{region 'Documentation'}
(*!
<summary>Check that IN is inside the inclusive StartTime..EndTime interval.</summary>
<description>

StartTime &gt; EndTime reports Error during active evaluation; equal bounds are
valid.

A value at or beyond 24 hours reports Error before comparison or baseline capture.

</description>
*)
{endregion}
FUNCTION_BLOCK AssertInTimespan_TOD EXTENDS AssertionBase
VAR_INPUT
    IN : TOD; //! Actual value checked or observed by this Assertion.
    StartTime : TOD; //! Inclusive start of the time span; must not exceed EndTime.
    EndTime : TOD; //! Inclusive end of the time span; must not precede StartTime.
END_VAR

SUPER^();

{region 'Documentation'}
(*!
<summary>Evaluate the typed temporal relation and report higher-priority errors first.</summary>
*)
{endregion}
METHOD PROTECTED Assert
VAR
    Message : STRING(GVL_Constants.MessageLength);
    StartTimeText : STRING(GVL_Constants.AssertionValueLength);
    EndTimeText : STRING(GVL_Constants.AssertionValueLength);
    ActualText : STRING(GVL_Constants.AssertionValueLength);
END_VAR
IF NOT EvaluationActive THEN
    RETURN;
END_IF;

IF Result = E_Result.Error THEN
    RETURN;
END_IF;

IF NOT IsTimeOfDayValid_TOD(Value := IN) THEN
    Error(Message := 'Assertion error: IN is outside the valid TOD range (less than 24 hours).');
    RETURN;
END_IF;

IF NOT IsTimeOfDayValid_TOD(Value := StartTime) THEN
    Error(Message := 'Assertion error: StartTime is outside the valid TOD range (less than 24 hours).');
    RETURN;
END_IF;

IF NOT IsTimeOfDayValid_TOD(Value := EndTime) THEN
    Error(Message := 'Assertion error: EndTime is outside the valid TOD range (less than 24 hours).');
    RETURN;
END_IF;

IF StartTime > EndTime THEN
    StartTimeText := TOD_TO_STRING(StartTime);
    EndTimeText := TOD_TO_STRING(EndTime);
    Message := CONCAT('Assertion error: start time exceeds end time. StartTime = ',
        StartTimeText);
    Message := CONCAT(Message, ', EndTime = ');
    Message := CONCAT(Message, EndTimeText);
    Message := CONCAT(Message, '.');
    Error(Message := Message);
    RETURN;
END_IF;

IF Result = E_Result.Failed THEN
    RETURN;
END_IF;

IF (IN < StartTime) OR (IN > EndTime) THEN
    StartTimeText := TOD_TO_STRING(StartTime);
    EndTimeText := TOD_TO_STRING(EndTime);
    ActualText := TOD_TO_STRING(IN);
    Message := CONCAT('Assertion failed: value is outside allowed timespan. StartTime = ',
        StartTimeText);
    Message := CONCAT(Message, ', EndTime = ');
    Message := CONCAT(Message, EndTimeText);
    Message := CONCAT(Message, ', Actual = ');
    Message := CONCAT(Message, ActualText);
    Message := CONCAT(Message, '.');
    Fail(Message := Message);
    RETURN;
END_IF;

Pass();
END_METHOD

END_FUNCTION_BLOCK

(* stored: Version 1.1.0.1
   POU AssertInTimespan_TOD: Id {4477cfb2-6d3f-4c5f-9156-77326181cd81}, SpecialFunc None
   Folder Internal: Id {2fa18933-22e7-479b-9910-39024a032ebe}
   Method Assert: Id {656454f8-f3bd-440e-9f74-63943618c596} *)
